Staubli VAL3: receive.pgx

public program receive()
  local bool l_bAckAlarm
  local bool l_bEndCmd
  local bool l_bErr
  local bool l_bHoldCmd
  local bool l_bPowerOff
  local bool l_bPowerOn
  local bool l_bResetCmd
  local bool l_bResetIO
  local bool l_bResult
  local bool l_bRotToHome
  local bool l_bStartCmd
  local bool l_bStopCmd
  local bool l_bToHome
  local bool l_bValue
  local num l_n
  local num l_nResult
  local num l_nSpeed
begin
  //机器人上电
  if dInPowerON==true and !isPowered() and workingMode()==4 and !rs:bIsEstop
    enablePower()
    l_bResult=watch(isPowered()==true,1)
    if !l_bResult
      popUpMsg("机器人上电超时")
    endIf
  endIf

  if rs:bIsCycle and workingMode()==1
    call cycle_stop()
  endIf
  //启动主程序
  if dInStartCycle==true and !rs:bIsCycle and rs:bIsHome and workingMode()==4 and !rs:bIsEstop
    //复位信号
    // call resetOutput()
    //
    //call cycle_stop()
    resetMotion()
    call cycle_start()
  endIf
  //暂停&恢复
  if dInPLCError==true
    if dOutGunON==true
      bSetGun=true
      dOutGunON=false
    endIf
    if rs:bIsCycle
      call cycle_pause()
    endIf
  elseIf dInPLCError==false and rs:bIsPause
    if bSetGun
      dOutGunON=true
    endIf
    call cycle_start()
  endIf
  //复位报警
  if dInResetError==true
    rs:bIsError=false
  endIf

  //设置速度
  call setSpeed()

  if esStatus()==1
    setSafetyRestart()
  endIf


end
